# B&R Automation Studio project POMiRTS_lab1
Automation Studio 4.5.2.102

## Configuration Config2

CPU 4PP065.0571-P74, AutomationRuntime D4.52, Build 4.1.2, Vc V4.52.0

### Task classes (Cpu.sw)
```
Cyclic#1:
  Program <- Program.prg
Binaries: udbdef, TCData, iomap, ashwac, Role, sysconf, arconfig, asfw, User, ashwd
Libraries: MotorContr
```

### Hardware
```
4PP065_0571_P74 : 4PP065.0571-P74 v1.1.2.0
  Connector IF5:
    ActivateDevice = 1
    Mode = Manual
    InternetAddress = 10.0.1.10
    SubnetMask = 255.255.255.0
  ConfigurationID = labBR
```

- Physical/Config2/4PP065_0571_P74/IoMap.iom: same as Physical/Config2/4PP065_0571_P74/Cpu.per
- Physical/Config2/4PP065_0571_P74/PvMap.vvm: same as Physical/Config2/4PP065_0571_P74/Cpu.per
## Logical view

Binary libraries used (declarations not repeated): operator, runtime, astime, AsIecCon

### Package Logical/Libraries - Global libraries

### Library Logical/Libraries/MotorContr (ANSIC)

#### MotorContr.fun - Exported functions and function blocks
```iecst
{REDUND_ERROR} {REDUND_UNREPLICABLE} FUNCTION_BLOCK FB_Integrator (*TODO: Add your comment here*) (*$GROUP=User,$CAT=User,$GROUPICON=User.png,$CATICON=User.png*)
	VAR_INPUT
		in : {REDUND_UNREPLICABLE} REAL;
	END_VAR
	VAR_OUTPUT
		out : {REDUND_UNREPLICABLE} REAL;
	END_VAR
	VAR
		dt : {REDUND_UNREPLICABLE} REAL;
	END_VAR
END_FUNCTION_BLOCK

{REDUND_ERROR} {REDUND_UNREPLICABLE} FUNCTION_BLOCK FB_Motor (*TODO: Add your comment here*) (*$GROUP=User,$CAT=User,$GROUPICON=User.png,$CATICON=User.png*)
	VAR_INPUT
		u : {REDUND_UNREPLICABLE} REAL;
	END_VAR
	VAR_OUTPUT
		w : {REDUND_UNREPLICABLE} REAL;
		phi : {REDUND_UNREPLICABLE} REAL;
	END_VAR
	VAR
		integrator : {REDUND_UNREPLICABLE} FB_Integrator;
		Tm : {REDUND_UNREPLICABLE} REAL;
		ke : {REDUND_UNREPLICABLE} REAL;
		dt : {REDUND_UNREPLICABLE} REAL;
	END_VAR
END_FUNCTION_BLOCK

{REDUND_ERROR} {REDUND_UNREPLICABLE} FUNCTION_BLOCK FB_Regulator (*TODO: Add your comment here*) (*$GROUP=User,$CAT=User,$GROUPICON=User.png,$CATICON=User.png*)
	VAR_INPUT
		e : {REDUND_UNREPLICABLE} REAL;
	END_VAR
	VAR_OUTPUT
		u : {REDUND_UNREPLICABLE} REAL;
	END_VAR
	VAR
		k_p : {REDUND_UNREPLICABLE} REAL;
		k_i : {REDUND_UNREPLICABLE} REAL;
		integrator : {REDUND_UNREPLICABLE} FB_Integrator;
		iyOld : {REDUND_UNREPLICABLE} REAL;
		max_abs_value : {REDUND_UNREPLICABLE} REAL;
		dt : {REDUND_UNREPLICABLE} REAL;
	END_VAR
END_FUNCTION_BLOCK
```

#### FB_Integrator.c
```c
#include <bur/plctypes.h>
#ifdef __cplusplus
	extern "C"
	{
#endif
	#include "MotorContr.h"
#ifdef __cplusplus
	};
#endif
/* TODO: Add your comment here */
void FB_Integrator(struct FB_Integrator* inst)
{
	inst->out = inst->in * inst->dt + inst->out;
}
```

#### FB_Motor.c
```c
#include <bur/plctypes.h>
#ifdef __cplusplus
	extern "C"
	{
#endif
	#include "MotorContr.h"
#ifdef __cplusplus
	};
#endif
/* TODO: Add your comment here */
void FB_Motor(struct FB_Motor* inst)
{
	/*TODO: Add your code here*/
	inst->w = (inst->u / inst->ke - inst->w) * (inst->dt / inst->Tm) + inst->w;
	inst->integrator.in = inst->w * 3.1415f / 30.0f; // С переводом в [рад/с]
	inst->integrator.dt = inst->dt;
	FB_Integrator(&inst->integrator);
	inst->phi = inst->integrator.out;
}
```

#### FB_Regulator.c
```c
ЫЫ#include <bur/plctypes.h>
#ifdef __cplusplus
	extern "C"
	{
#endif
	#include "MotorContr.h"
#ifdef __cplusplus
	};
#endif
/* TODO: Add your comment here */
void FB_Regulator(struct FB_Regulator* inst)
{
	/*TODO: Add your code here*/
	float proportial = inst->e * inst->k_p;
	if (proportial > inst->max_abs_value)
	{
		proportial = inst->max_abs_value;
	}
	else if ( proportial < -inst->max_abs_value)
	{
		proportial = -inst->max_abs_value;
	}
	float integral_part_in = inst->e * inst->k_i - inst->iyOld / inst->dt;
	inst->integrator.in = integral_part_in;
	inst->integrator.dt = inst->dt;
	FB_Integrator(&inst->integrator);
	float sum = proportial + inst->integrator.out;

	if (sum > inst->max_abs_value)
	{
		inst->u = inst->max_abs_value;
	}
	else if (sum < -inst->max_abs_value)
	{
		inst->u = -inst->max_abs_value;
	}
	else inst->u = sum;

	inst->iyOld = sum - inst->u;
}
```

### Program Logical/Program (ANSIC)

#### Main.c - Init, cyclic, exit code
```c
#include <bur/plctypes.h>
#ifdef _DEFAULT_INCLUDES
	#include <AsDefault.h>
#endif

void _INIT ProgramInit(void)
{
	fb_regulator.dt = 0.01f;
	fb_motor.dt = 0.01f;
	fb_motor2.dt = 0.01f;
	fb_motor.ke = 0.02f;
	fb_motor.Tm = 0.08f;
	fb_motor2.ke = 0.002f;
	fb_motor2.Tm = 0.08f;
	fb_regulator.max_abs_value = 50;
	fb_regulator.k_i = 0.80f;
	fb_regulator.k_p = 0.16f;
	fb_regulator.iyOld = 0.0f;

	fb_motor.w = 0.0f;
	fb_motor.integrator.out = 0.0f;
	fb_motor2.w = 0.0f;
	fb_motor2.integrator.out = 0.0f;
	counter = 0;
	speed = 0.0f;
	fb_regulator.integrator.out = 0.0f;
	Enable = 1;
}

void motor_regulated() {
	if (!Enable){
		fb_regulator.u = 0.0f;
		fb_regulator.iyOld = 0.0f;
		fb_regulator.integrator.out = 0.0f;
		fb_motor.u = 0.0f;
		FB_Motor(&fb_motor);
	}
	else{
		fb_regulator.e = speed - fb_motor.w;
		FB_Regulator(&fb_regulator);
		fb_motor.u = fb_regulator.u;
		FB_Motor(&fb_motor);
	}
}

void motor_unregulated() {
	if (!Enable) {
		fb_motor2.u = 0.0f;
		fb_motor2.w = 0.0f;
		fb_motor2.phi = 0.0f;
		FB_Motor(&fb_motor2);
		return;
	}
	else {
		fb_motor2.u = speed * fb_motor2.ke;
		FB_Motor(&fb_motor2);
	}
}

void stupench() {
	if (!Enable) {
		counter = 0;
		speed = 0.0f;
	}
	else{
		counter++;
		if (counter < 500)
			speed = 0.0f;
		else if (counter < 1000)
			speed = 800.0f;
		else {
			speed = 0.0f;
			counter = 0;
		}
	}
}

void _CYCLIC ProgramCyclic(void)
{
	stupench();
	motor_regulated();
	motor_unregulated();
}

void _EXIT ProgramExit(void)
{
}
```

#### Variables.var - Local variables
```iecst
VAR
	counter : INT := 0;
	fb_motor2 : FB_Motor;
	Enable : BOOL := TRUE;
	speed : REAL;
	fb_motor : FB_Motor;
	fb_regulator : FB_Regulator;
END_VAR
```
